// TIA Portal V20 export
// export: Created 2026-10-20T12:40:41.0438244Z, ExportSetting WithDefaults, DisplayName Totally Integrated Automation Portal, DisplayVersion V20 Update 6, DisplayName TIA Portal Openness, DisplayVersion V20 Update 6, DisplayName TIA Portal Version Control Interface, DisplayVersion V20 Update 6, DisplayName SINAMICS Startdrive Advanced, DisplayVersion V20 SP1, DisplayName SINAMICS Startdrive G130, G150, S120, S150, SINAMICS MV, G220, S200, S210, DisplayVersion V20 SP1, DisplayName SINAMICS Startdrive G110M, G120, G120C, G120D, G120P, G115D, DisplayVersion V20 SP1, DisplayName STEP 7 Professional, DisplayVersion V20 Update 6, DisplayName STEP 7 Safety, DisplayVersion V20 Update 2, DisplayName WinCC Basic/Comfort/Advanced, DisplayVersion V20 Update 6, DisplayName WinCC Unified, DisplayVersion V20 Update 6
FUNCTION "SICK_SetValue" : Void   // FC11, SCL
TITLE = Set value
{ S7_Optimized_Access := 'TRUE' }
AUTHOR : SICKAG
FAMILY : Ident
VERSION : 1.1
// This function is needs to set a value to a SICK CoLa command.
// stored: AutoNumber false, IsIECCheckEnabled false, SetENOAutomatically false, UDAEnableTagReadback false
   VAR_INPUT
      bAddBlank : Bool;   // Add blank after value
      nValue : DWord;   // Value that should be written
   END_VAR
   VAR_OUTPUT
      arrData : Array[0..499] of Byte;   // Destination telegram
      nErrorCode : Word;   // Error code
   END_VAR
   VAR_IN_OUT
      iPosition : UInt;   // Position offset of the value before and after (starting from 0)
   END_VAR
   VAR_TEMP
      iValueLength : USInt;   // Byte length of the value that shuld be written
      nReturnValue : Word;   // Return value of the convert function
      sValue : String[8];   // Converted value
      nTempValue : DWord;   // Temporarily variable
      iTemp : UInt;   // Temporarily variable
   END_VAR
BEGIN
   (*===========================================================================================
   Name:   SICK_SetValue
   Author: SICK AG
   =============================================================================================
   Description: 
   This function is for internal use only.
   The function converts a hexadecimal value into a hexadecimal string and add it 
   automatically to the command array.     

   =============================================================================================
   Error codes:
   16#0000 = No error
   16#0001 = Invalid position index   
   16#8xxx = Conversion error (HTA-Function) see help system for more information

   =============================================================================================
   Version history:
   Date       | Version | created under               | Author  | Remark
   ---------------------------------------------------------------------------------------------
   30/01/2014 | V1.0    | TIA Portal V12 SP1 Update 2 | SICK AG | Initial version
   22/04/2014 | V1.1    | TIA Portal V12 SP1 Update 4 | SICK AG | Avoid warnings that occur with 
                                                                  TIA V13
   ============================================================================================*)

   (*===================================== INITIALISATION =====================================*)
   #iValueLength:= 0;
   #nErrorCode:= 16#0000;

   (*======================================= WRITE VALUE ======================================*)
   (*Check current position of the value*)
   IF #iPosition > 499 THEN 
     #nErrorCode:= 16#0001; (*Error: Invalid position index*)
     RETURN;
   END_IF;



   (*Get byte length of the value that should be written*)
   IF #nValue <= 16#FF THEN
     #nTempValue:= SHL(IN:= #nValue, N:=24);
     #iValueLength:= 1;
   ELSIF #nValue <= 16#FFFF THEN
     #nTempValue:= SHL(IN:= #nValue, N:=16);
     #iValueLength:= 2;
   ELSIF #nValue <= 16#00FF_FFFF THEN
     #nTempValue:= SHL(IN:= #nValue, N:=8);
     #iValueLength:= 3;
   ELSIF #nValue <= 16#FFFF_FFFF THEN
     #nTempValue:= #nValue;
     #iValueLength:= 4;
   END_IF;

   (*Convert hexadecimal number into a ASCII string*)
   #nReturnValue:= HTA(IN:= #nTempValue, N:= #iValueLength, OUT=>#sValue);
   IF #nReturnValue <> 16#0000 THEN
     #nErrorCode:= #nReturnValue; (*Error: Conversion error (HTA-Function)*)
     RETURN;
   END_IF;

   (*Add the string value to the destination telegram*)
   #arrData[#iPosition]:= 0; // Avoid warnings under TIA V13
   Strg_TO_Chars(Strg:=#sValue, pChars:= #iPosition, Cnt=> #iTemp, Chars:= #arrData);

   (*Add blank to the destination telegram and calculate the position of the next element*)
   IF #bAddBlank THEN
     #arrData[#iPosition+#iTemp]:= ' ';
     #iPosition:= #iPosition+#iTemp+1;

   (*Calculate the position of the next element*)
   ELSE
     #iPosition:= #iPosition+#iTemp;
   END_IF;
END_FUNCTION
